(* IEC 61131-3 sources: Elmo_Master/Lasal_PRG/MotionTCPDemo/Network/TCPComNet, 1 file *)

(* ---- ONE_TCPComNet_Table.st ---- *)
#define OBJECTS_CONFIG

#include "..\..\Class\DataManager\DataManager.h"
//Define part of class DataManagerFIFO
#define MEMORY_Mark_DataMngFiFo    8
#include <.\lsl_st_mt.h>
#include "..\..\Class\TCPCommunication\TCPCommunication.h"
#include "..\..\Class\TCPCommunication\SalamanderDelay.h"

FUNCTION GLOBAL TAB ONE_TCPComNet
-1$UINT, 0$UINT,
0$UINT, 0$UINT,

17$UDINT,
TO_UDINT(916194998), "_CheckSum", 1$UINT, 0$UINT, 1$UINT,
TO_UDINT(3238142347), "_SigTCPComReceive", 1$UINT, 1$UINT, 0$UINT,
TO_UDINT(969826267), "_SigTCPDataManager", 1$UINT, 1$UINT, 0$UINT,
TO_UDINT(794617671), "CriticalSection", 0$UINT, 4$UINT, 10$UINT,
TO_UDINT(4008337867), "DataManager", 1$UINT, 1$UINT, 0$UINT,
TO_UDINT(2873804345), "DataManagerFIFO", 1$UINT, 1$UINT, 10$UINT,
TO_UDINT(2393054465), "DataManagerPriority", 1$UINT, 0$UINT, 1$UINT,
TO_UDINT(2602835227), "GetTaskHandle", 0$UINT, 2$UINT, 1$UINT,
TO_UDINT(2225119864), "MerkerEx", 1$UINT, 22$UINT, 2$UINT,
TO_UDINT(3534980377), "RamRingBuffer", 1$UINT, 1$UINT, 1$UINT,
TO_UDINT(1240328812), "ReceiveMsg", 0$UINT, 0$UINT, 1$UINT,
TO_UDINT(1850111279), "String", 1$UINT, 11$UINT, 1$UINT,
TO_UDINT(2898603620), "StringInternal", 1$UINT, 86$UINT, 0$UINT,
TO_UDINT(4051501096), "TCP_MotionIF_Dummy", 0$UINT, 0$UINT, 1$UINT,
TO_UDINT(3704218787), "TCPCommunication", 1$UINT, 20$UINT, 1$UINT,
TO_UDINT(3171666764), "TCPRT_DataManager", 0$UINT, 0$UINT, 1$UINT,
TO_UDINT(3232495061), "VirtualBaseInit", 1$UINT, 3$UINT, 0$UINT,

1$UINT, TO_UDINT(2771092362), "_SIGTCPDATAMANAGER1\_BASE\TCPCOMMUNICATION\CHECKSUM",

1$UINT, TO_UDINT(834118171), "_SIGTCPDATAMANAGER1\_BASE\_BASE\DATAMANAGERPRIORITY\DATAMANAGERFIFO_PRIO0\SECTION",
1$UINT, TO_UDINT(650950232), "_SIGTCPDATAMANAGER1\_BASE\_BASE\DATAMANAGERPRIORITY\DATAMANAGERFIFO_PRIO1\SECTION",
1$UINT, TO_UDINT(524389021), "_SIGTCPDATAMANAGER1\_BASE\_BASE\DATAMANAGERPRIORITY\DATAMANAGERFIFO_PRIO2\SECTION",
1$UINT, TO_UDINT(138059486), "_SIGTCPDATAMANAGER1\_BASE\_BASE\DATAMANAGERPRIORITY\DATAMANAGERFIFO_PRIO3\SECTION",
1$UINT, TO_UDINT(1817965335), "_SIGTCPDATAMANAGER1\_BASE\_BASE\DATAMANAGERPRIORITY\DATAMANAGERFIFO_PRIO4\SECTION",
1$UINT, TO_UDINT(2065753940), "_SIGTCPDATAMANAGER1\_BASE\_BASE\DATAMANAGERPRIORITY\DATAMANAGERFIFO_PRIO5\SECTION",
1$UINT, TO_UDINT(1118690193), "_SIGTCPDATAMANAGER1\_BASE\_BASE\DATAMANAGERPRIORITY\DATAMANAGERFIFO_PRIO6\SECTION",
1$UINT, TO_UDINT(1440141266), "_SIGTCPDATAMANAGER1\_BASE\_BASE\DATAMANAGERPRIORITY\DATAMANAGERFIFO_PRIO7\SECTION",
1$UINT, TO_UDINT(2322530307), "_SIGTCPDATAMANAGER1\_BASE\_BASE\DATAMANAGERPRIORITY\DATAMANAGERFIFO_PRIO8\SECTION",
1$UINT, TO_UDINT(2635338816), "_SIGTCPDATAMANAGER1\_BASE\_BASE\DATAMANAGERPRIORITY\DATAMANAGERFIFO_PRIO9\SECTION",

1$UINT, TO_UDINT(2700156713), "_SIGTCPDATAMANAGER1\_BASE\_BASE\DATAMANAGERPRIORITY\DATAMANAGERFIFO_PRIO0",
1$UINT, TO_UDINT(3623235519), "_SIGTCPDATAMANAGER1\_BASE\_BASE\DATAMANAGERPRIORITY\DATAMANAGERFIFO_PRIO1",
1$UINT, TO_UDINT(1325366789), "_SIGTCPDATAMANAGER1\_BASE\_BASE\DATAMANAGERPRIORITY\DATAMANAGERFIFO_PRIO2",
1$UINT, TO_UDINT(972574355), "_SIGTCPDATAMANAGER1\_BASE\_BASE\DATAMANAGERPRIORITY\DATAMANAGERFIFO_PRIO3",
1$UINT, TO_UDINT(2812074800), "_SIGTCPDATAMANAGER1\_BASE\_BASE\DATAMANAGERPRIORITY\DATAMANAGERFIFO_PRIO4",
1$UINT, TO_UDINT(3499879334), "_SIGTCPDATAMANAGER1\_BASE\_BASE\DATAMANAGERPRIORITY\DATAMANAGERFIFO_PRIO5",
1$UINT, TO_UDINT(1234352668), "_SIGTCPDATAMANAGER1\_BASE\_BASE\DATAMANAGERPRIORITY\DATAMANAGERFIFO_PRIO6",
1$UINT, TO_UDINT(1049987722), "_SIGTCPDATAMANAGER1\_BASE\_BASE\DATAMANAGERPRIORITY\DATAMANAGERFIFO_PRIO7",
1$UINT, TO_UDINT(2922026779), "_SIGTCPDATAMANAGER1\_BASE\_BASE\DATAMANAGERPRIORITY\DATAMANAGERFIFO_PRIO8",
1$UINT, TO_UDINT(3643647885), "_SIGTCPDATAMANAGER1\_BASE\_BASE\DATAMANAGERPRIORITY\DATAMANAGERFIFO_PRIO9",

1$UINT, TO_UDINT(3030441658), "_SIGTCPDATAMANAGER1\_BASE\_BASE\DATAMANAGERPRIORITY",

1$UINT, TO_UDINT(3628408059), "_SIGTCPDATAMANAGER1\_BASE\_BASE\DATAMNGGETTASKHANDLE1",

1$UINT, TO_UDINT(552288716), "_SIGTCPDATAMANAGER1\_BASE\TCPCOMMUNICATION\RAMRINGMERKEREX",
1$UINT, TO_UDINT(285254243), "_SIGTCPDATAMANAGER1\_BASE\TCPCOMMUNICATION\THREADNAME\MERKEREX0",

1$UINT, TO_UDINT(1506338805), "_SIGTCPDATAMANAGER1\_BASE\TCPCOMMUNICATION\RAMRINGBUFFER",

_NO_ATTR, TO_UDINT(3348180782), "RECEIVEMSG1",

1$UINT, TO_UDINT(2598389583), "_SIGTCPDATAMANAGER1\_BASE\TCPCOMMUNICATION\THREADNAME",

_NO_ATTR, TO_UDINT(3063429709), "TCP_MOTIONIF_DUMMY1",

1$UINT, TO_UDINT(3493563493), "_SIGTCPDATAMANAGER1\_BASE\TCPCOMMUNICATION",

_NO_ATTR, TO_UDINT(2464426676), "_SIGTCPDATAMANAGER1",

//Internal connections
0$UDINT,
28$UDINT,
TO_UDINT(11), "Section", TO_UDINT(1),
TO_UDINT(12), "Section", TO_UDINT(2),
TO_UDINT(13), "Section", TO_UDINT(3),
TO_UDINT(14), "Section", TO_UDINT(4),
TO_UDINT(15), "Section", TO_UDINT(5),
TO_UDINT(16), "Section", TO_UDINT(6),
TO_UDINT(17), "Section", TO_UDINT(7),
TO_UDINT(18), "Section", TO_UDINT(8),
TO_UDINT(19), "Section", TO_UDINT(9),
TO_UDINT(20), "Section", TO_UDINT(10),
TO_UDINT(21), "DataManagerFiFo_Prio0", TO_UDINT(11),
TO_UDINT(21), "DataManagerFiFo_Prio1", TO_UDINT(12),
TO_UDINT(21), "DataManagerFiFo_Prio2", TO_UDINT(13),
TO_UDINT(21), "DataManagerFiFo_Prio3", TO_UDINT(14),
TO_UDINT(21), "DataManagerFiFo_Prio4", TO_UDINT(15),
TO_UDINT(21), "DataManagerFiFo_Prio5", TO_UDINT(16),
TO_UDINT(21), "DataManagerFiFo_Prio6", TO_UDINT(17),
TO_UDINT(21), "DataManagerFiFo_Prio7", TO_UDINT(18),
TO_UDINT(21), "DataManagerFiFo_Prio8", TO_UDINT(19),
TO_UDINT(21), "DataManagerFiFo_Prio9", TO_UDINT(20),
TO_UDINT(27), "MerkerEx0", TO_UDINT(24),
TO_UDINT(29), "RamRingBuffer", TO_UDINT(25),
TO_UDINT(29), "RamRingMerkerEx", TO_UDINT(23),
TO_UDINT(29), "CheckSum", TO_UDINT(0),
TO_UDINT(29), "ThreadName", TO_UDINT(27),
TO_UDINT(30), "DataMngGetTaskHandle1", TO_UDINT(22),
TO_UDINT(30), "DataManagerPriority", TO_UDINT(21),
TO_UDINT(30), "TCPCommunication", TO_UDINT(29),
0$UDINT,
6$UDINT,
TO_UDINT(25), "Data", TO_UDINT(23), "m_udLength",
TO_UDINT(26), "_SigTCPDataManager", TO_UDINT(30), "ClassSvr",
TO_UDINT(27), "DataBuffer", TO_UDINT(24), "m_udLength",
TO_UDINT(28), "_SigTCPDataManager", TO_UDINT(30), "ClassSvr",
TO_UDINT(29), "coDataMng", TO_UDINT(30), "ClassSvr",
TO_UDINT(30), "coTCPCommunication", TO_UDINT(29), "ClassSvr",

//Initialization values
0$UDINT,
18$UDINT,
TO_UDINT(23), "ThreadSafe", TO_UDINT(0),//|TCPComNet.TCPCommunication\_base\_SigTCPDataManager1\RamRingMerkerEx.ThreadSafe;
TO_UDINT(24), "ThreadSafe", TO_UDINT(0),//|TCPComNet.ThreadName\TCPCommunication\_base\_SigTCPDataManager1\MerkerEx0.ThreadSafe;
TO_UDINT(26), "SourceID", TO_UDINT(101),//|TCPComNet.ReceiveMsg1.SourceID;
TO_UDINT(27), "SingleRealloc", TO_UDINT(1),//|TCPComNet.TCPCommunication\_base\_SigTCPDataManager1\ThreadName.SingleRealloc;
TO_UDINT(28), "SourceID", TO_UDINT(1),//|TCPComNet.TCP_MotionIF_Dummy1.SourceID;
TO_UDINT(29), "ComPort", TO_UDINT(500),//|TCPComNet._base\_SigTCPDataManager1\TCPCommunication.ComPort;
TO_UDINT(29), "LogEnable", TO_UDINT(0),//|TCPComNet._base\_SigTCPDataManager1\TCPCommunication.LogEnable;
TO_UDINT(29), "DeactivateCom", TO_UDINT(0),//|TCPComNet._base\_SigTCPDataManager1\TCPCommunication.DeactivateCom;
TO_UDINT(29), "coLogFilter", TO_UDINT(0),//|TCPComNet._base\_SigTCPDataManager1\TCPCommunication.coLogFilter;
TO_UDINT(29), "SizeOfComBuffers", TO_UDINT(100 kB),//|TCPComNet._base\_SigTCPDataManager1\TCPCommunication.SizeOfComBuffers;
TO_UDINT(29), "SizeOfComBufferRecv", TO_UDINT(100 kB),//|TCPComNet._base\_SigTCPDataManager1\TCPCommunication.SizeOfComBufferRecv;
TO_UDINT(30), "AcceptOfflineJobs", TO_UDINT(1),//|TCPComNet._SigTCPDataManager1.AcceptOfflineJobs;
TO_UDINT(30), "ComPort", TO_UDINT(500),//|TCPComNet._SigTCPDataManager1.ComPort;
TO_UDINT(30), "LogEnable", TO_UDINT(0),//|TCPComNet._SigTCPDataManager1.LogEnable;
TO_UDINT(30), "DeactivateCom", TO_UDINT(0),//|TCPComNet._SigTCPDataManager1.DeactivateCom;
TO_UDINT(30), "LogFilter", TO_UDINT(0),//|TCPComNet._SigTCPDataManager1.LogFilter;
TO_UDINT(30), "SizeOfComBuffers", TO_UDINT(100 kB),//|TCPComNet._SigTCPDataManager1.SizeOfComBuffers;
TO_UDINT(30), "SizeOfComBufferRecv", TO_UDINT(100 kB),//|TCPComNet._SigTCPDataManager1.SizeOfComBufferRecv;

//Symbolic initialization values
0$UDINT,
0$UDINT,

//Initialization of string values
0$UDINT,
0$UDINT,

//Configuration of tasks (RealTime, Cyclic, Background)
0$UDINT,
1$UDINT,
TO_UDINT(22), (1000)$UDINT, 4194303$DINT, 	//_SIGTCPDATAMANAGER1\_BASE\_BASE\DATAMNGGETTASKHANDLE1

0$UDINT,
1$UDINT,
TO_UDINT(22), (1000)$UDINT, 4194303$DINT, 	//_SIGTCPDATAMANAGER1\_BASE\_BASE\DATAMNGGETTASKHANDLE1

0$UDINT,
1$UDINT,
TO_UDINT(22), (1000)$UDINT, 4194303$DINT, 	//_SIGTCPDATAMANAGER1\_BASE\_BASE\DATAMNGGETTASKHANDLE1

//External connections
0$UDINT,
0$UDINT,

//Magic internal connections
0$UDINT,
7$UDINT,
TO_UDINT(29), "coIntern", TO_UDINT(30), "InternConnection",
TO_UDINT(29), "coIpToConnect", TO_UDINT(30), "IPtoConnect",
TO_UDINT(29), "coStationToConnect", TO_UDINT(30), "StationToConnect",
TO_UDINT(29), "coLogFilter", TO_UDINT(30), "LogFilter",
TO_UDINT(29), "ErrRuntime", TO_UDINT(30), "ErrRuntime",
TO_UDINT(29), "SizeOfComBuffers", TO_UDINT(30), "SizeOfComBuffers",
TO_UDINT(29), "SizeOfComBufferRecv", TO_UDINT(30), "SizeOfComBufferRecv",

//Configuration of timeslots of tasks (RealTime, Cyclic)
#ifdef __LSLLDR_TIMESLOTS__
0$UDINT,
0$UDINT,

0$UDINT,
0$UDINT,

#endif //__LSLLDR_TIMESLOTS__

//MultiMaster connections
#ifdef __LSLLDR_MULTIMASTER__
0$UDINT,
0$UDINT,
#endif //__LSLLDR_MULTIMASTER__

//Configuration for task ID (RealTime, CyclicTime)
#ifdef __LSLLDR_TASKID__
"\\\\TASKS2  "
0$UDINT,
1$UDINT,
(0)$UDINT, 	//_SIGTCPDATAMANAGER1\_BASE\_BASE\DATAMNGGETTASKHANDLE1

0$UDINT,
1$UDINT,
(0)$UDINT, 	//_SIGTCPDATAMANAGER1\_BASE\_BASE\DATAMNGGETTASKHANDLE1

0$UDINT,
1$UDINT,
(0)$UDINT, 	//_SIGTCPDATAMANAGER1\_BASE\_BASE\DATAMNGGETTASKHANDLE1

#endif //__LSLLDR_TASKID__

END_FUNCTION
